DATA_BLOCK "FRK_HostStore"
{ S7_Optimized_Access := 'TRUE' }
VERSION : 0.1
NON_RETAIN
VAR
    Rows {ExternalAccessible := 'False'; ExternalVisible := 'False'; ExternalWritable := 'False'} : Array[1..1] of "FRK_HostBook";
END_VAR
BEGIN
END_DATA_BLOCK
